// CFC twin of T_SafeTwoHand_Tests: the same tests drawn as CFC diagrams, the way a TwinSAFE project is authored.
    FUNCTION_BLOCK T_SafeTwoHand_Tests_CFC EXTENDS T_SafeCfcTestSuite
    VAR
    // Test_BothHandsGiveOutputAndReleaseNeedsBothOff
    group_1 : T_SafeGroup;
    fb_1 : T_SafeTwoHand(group := group_1);
    // Test_SecondHandWithoutFirstGivesTwoHandError
    group_2 : T_SafeGroup;
    fb_2 : T_SafeTwoHand(group := group_2);
    // Test_HandDiscrepancyTimeout
    group_3 : T_SafeGroup;
    // SafeInputsAfterDiscError TRUE (not the default) so the error waits for both hands released (diag bit 10)
    fb_3 : T_SafeTwoHand(group := group_3) := (Parameters := (HandDiscrepancyTime := T#100MS, SafeInputsAfterDiscError := TRUE));
    t0_3 : TON;
    t1_3 : TON;
    trig1_3 : R_TRIG;
END_VAR

Test_BothHandsGiveOutputAndReleaseNeedsBothOff();
Test_SecondHandWithoutFirstGivesTwoHandError();
Test_HandDiscrepancyTimeout();

METHOD PRIVATE Test_BothHandsGiveOutputAndReleaseNeedsBothOff
// note: this text did not pass the execution check against the stored diagram
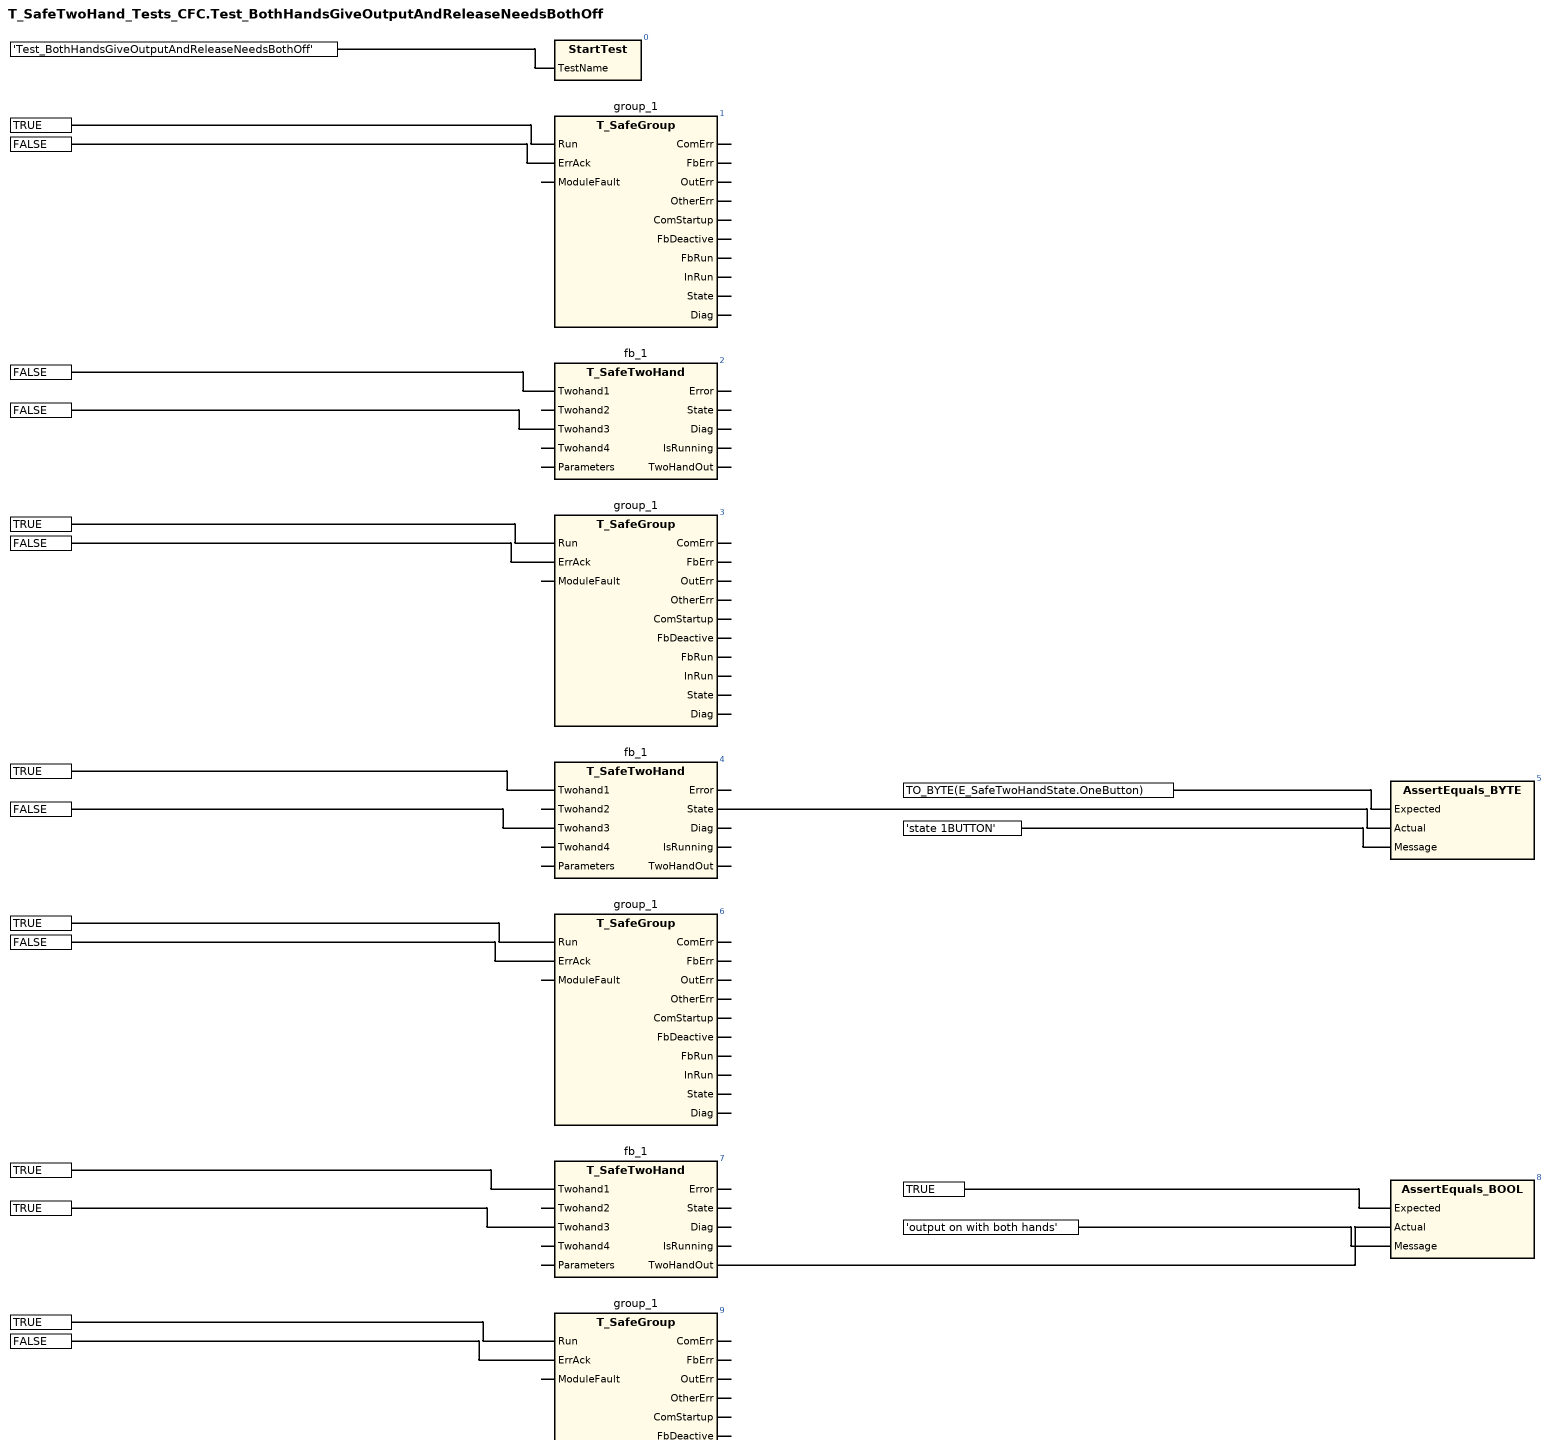
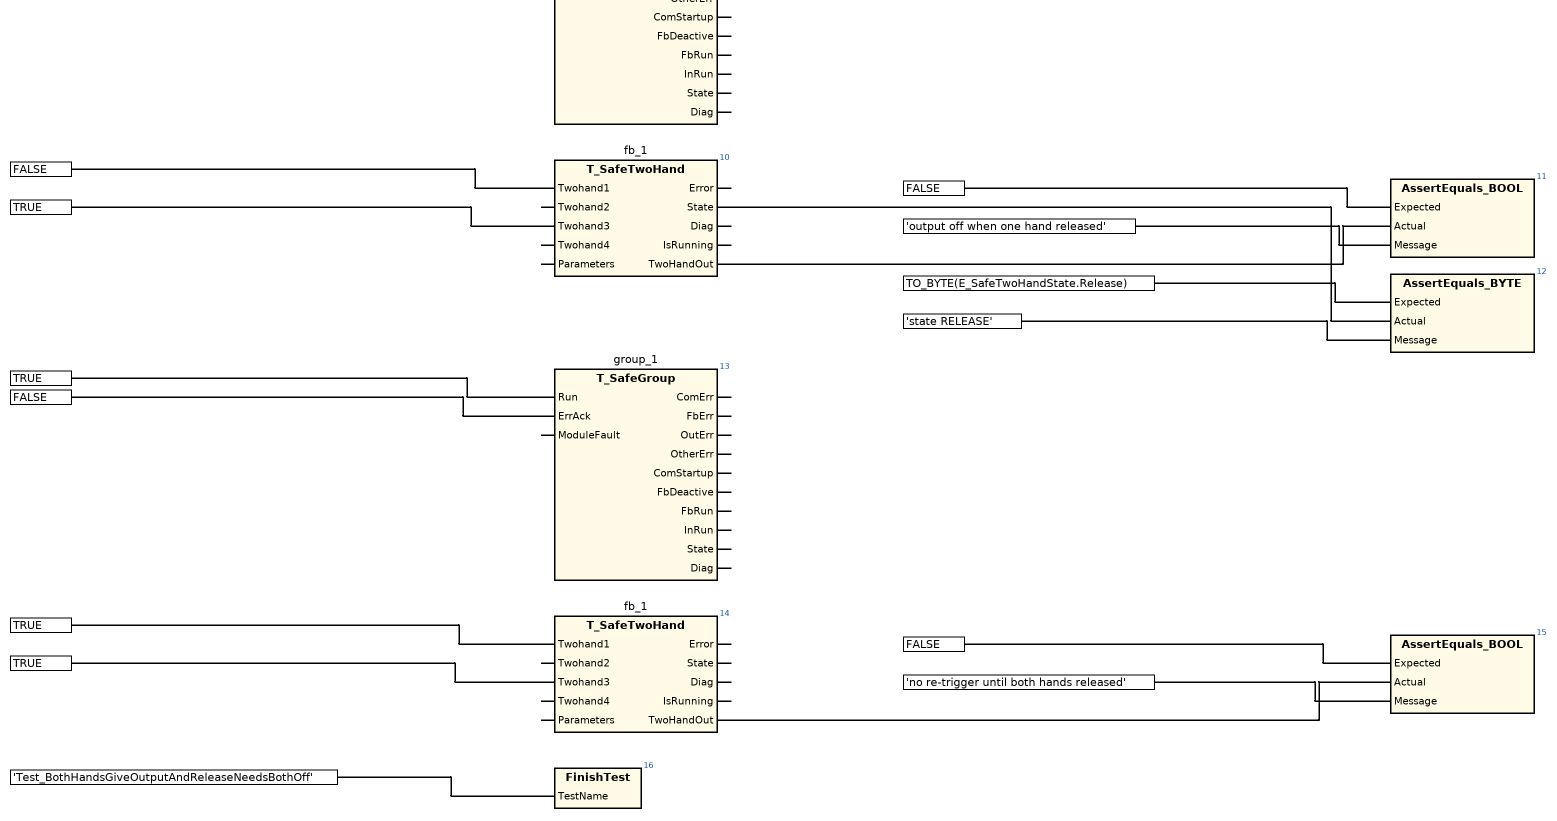
StartTest(TestName := 'Test_BothHandsGiveOutputAndReleaseNeedsBothOff');
group_1(Run := TRUE, ErrAck := FALSE); // T_SafeGroup
fb_1(Twohand1 := FALSE, Twohand3 := FALSE); // T_SafeTwoHand
group_1(Run := TRUE, ErrAck := FALSE); // T_SafeGroup
fb_1(Twohand1 := TRUE, Twohand3 := FALSE); // T_SafeTwoHand
AssertEquals_BYTE(Expected := TO_BYTE(E_SafeTwoHandState.OneButton), Actual := fb_1.State, Message := 'state 1BUTTON');
group_1(Run := TRUE, ErrAck := FALSE); // T_SafeGroup
fb_1(Twohand1 := TRUE, Twohand3 := TRUE); // T_SafeTwoHand
AssertEquals_BOOL(Expected := TRUE, Actual := fb_1.TwoHandOut, Message := 'output on with both hands');
group_1(Run := TRUE, ErrAck := FALSE); // T_SafeGroup
fb_1(Twohand1 := FALSE, Twohand3 := TRUE); // T_SafeTwoHand
AssertEquals_BOOL(Expected := FALSE, Actual := fb_1.TwoHandOut, Message := 'output off when one hand released');
AssertEquals_BYTE(Expected := TO_BYTE(E_SafeTwoHandState.Release), Actual := fb_1.State, Message := 'state RELEASE');
group_1(Run := TRUE, ErrAck := FALSE); // T_SafeGroup
fb_1(Twohand1 := TRUE, Twohand3 := TRUE); // T_SafeTwoHand
AssertEquals_BOOL(Expected := FALSE, Actual := fb_1.TwoHandOut, Message := 'no re-trigger until both hands released');
FinishTest(TestName := 'Test_BothHandsGiveOutputAndReleaseNeedsBothOff');
END_METHOD

METHOD PRIVATE Test_SecondHandWithoutFirstGivesTwoHandError
// note: this text did not pass the execution check against the stored diagram
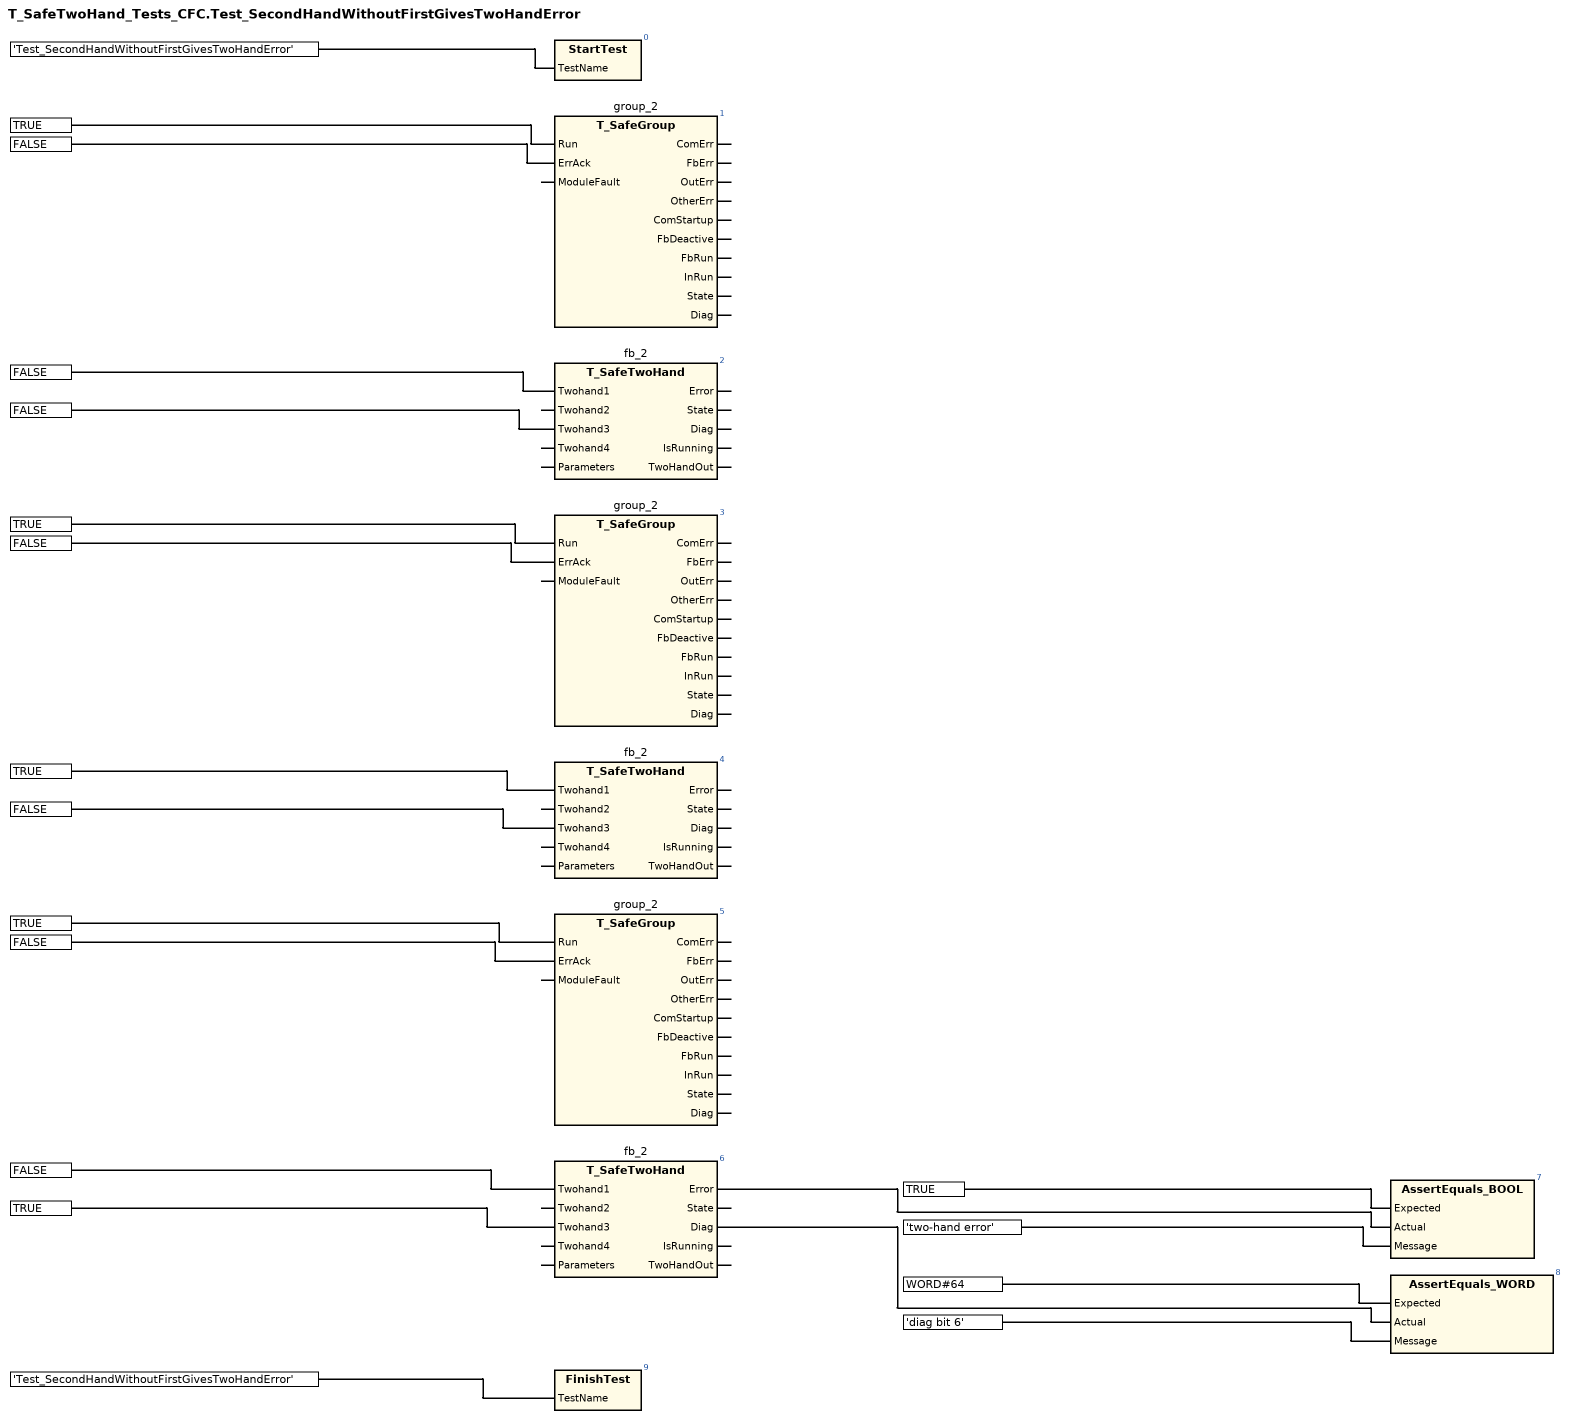
StartTest(TestName := 'Test_SecondHandWithoutFirstGivesTwoHandError');
group_2(Run := TRUE, ErrAck := FALSE); // T_SafeGroup
fb_2(Twohand1 := FALSE, Twohand3 := FALSE); // T_SafeTwoHand
group_2(Run := TRUE, ErrAck := FALSE); // T_SafeGroup
fb_2(Twohand1 := TRUE, Twohand3 := FALSE); // T_SafeTwoHand
group_2(Run := TRUE, ErrAck := FALSE); // T_SafeGroup
fb_2(Twohand1 := FALSE, Twohand3 := TRUE); // T_SafeTwoHand
AssertEquals_BOOL(Expected := TRUE, Actual := fb_2.Error, Message := 'two-hand error');
AssertEquals_WORD(Expected := WORD#64, Actual := fb_2.Diag, Message := 'diag bit 6');
FinishTest(TestName := 'Test_SecondHandWithoutFirstGivesTwoHandError');
END_METHOD

METHOD PRIVATE Test_HandDiscrepancyTimeout
// note: this text did not pass the execution check against the stored diagram
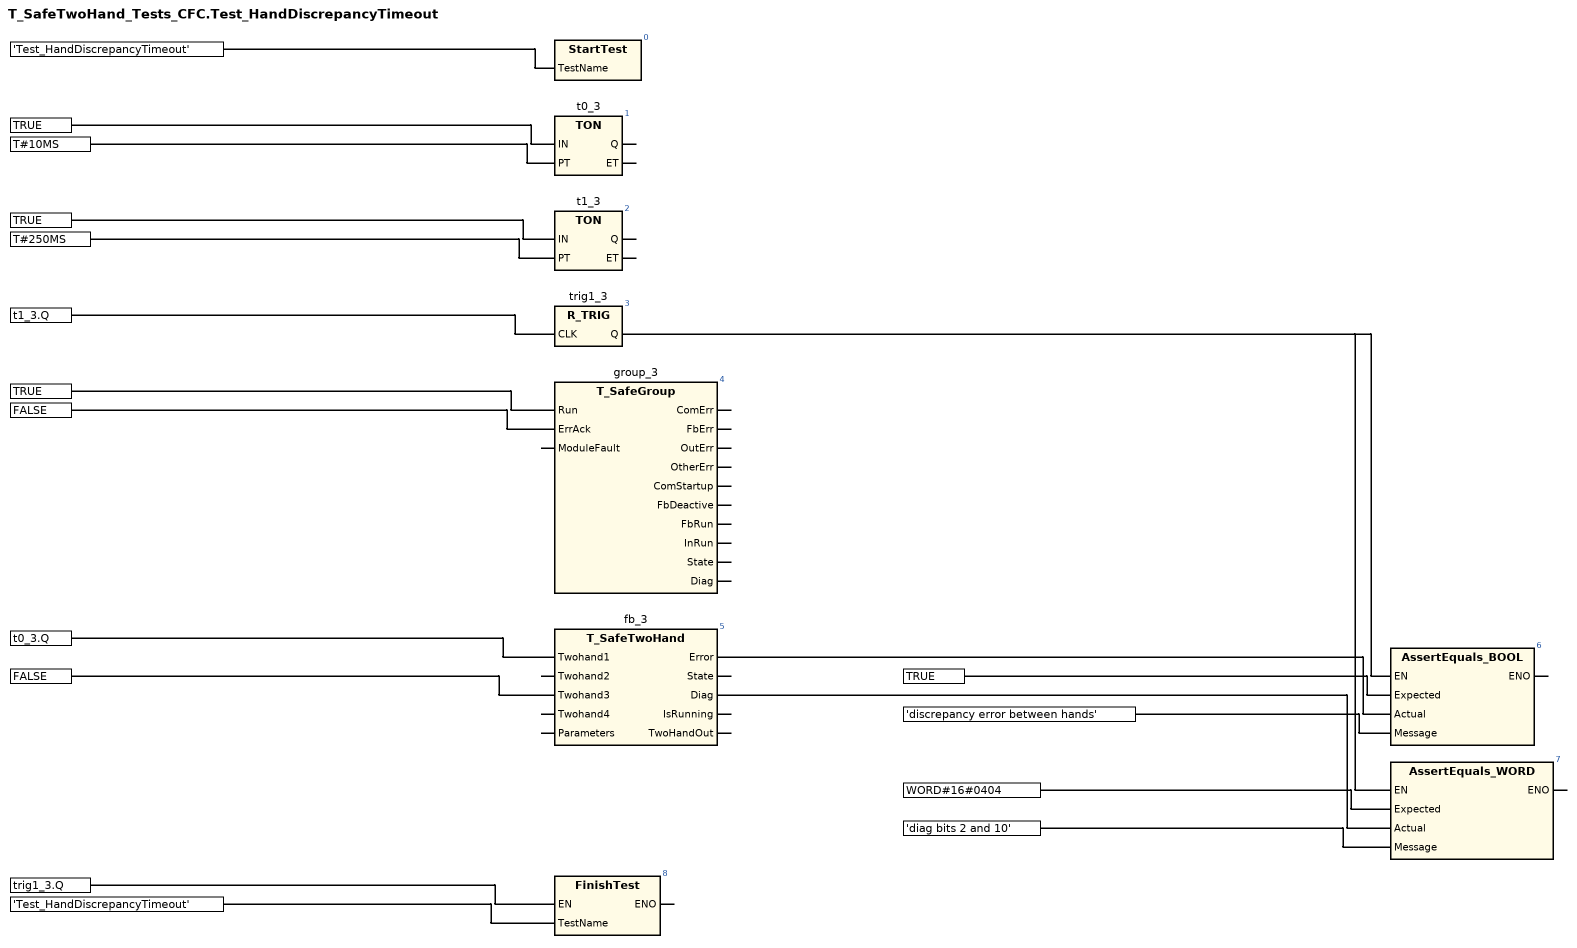
StartTest(TestName := 'Test_HandDiscrepancyTimeout');
t0_3(IN := TRUE, PT := T#10MS); // TON
t1_3(IN := TRUE, PT := T#250MS); // TON
trig1_3(CLK := t1_3.Q); // R_TRIG
group_3(Run := TRUE, ErrAck := FALSE); // T_SafeGroup
fb_3(Twohand1 := t0_3.Q, Twohand3 := FALSE); // T_SafeTwoHand
IF trig1_3.Q THEN AssertEquals_BOOL(Expected := TRUE, Actual := fb_3.Error, Message := 'discrepancy error between hands'); END_IF
IF trig1_3.Q THEN AssertEquals_WORD(Expected := WORD#16#0404, Actual := fb_3.Diag, Message := 'diag bits 2 and 10'); END_IF
IF trig1_3.Q THEN FinishTest(TestName := 'Test_HandDiscrepancyTimeout'); END_IF
END_METHOD

END_FUNCTION_BLOCK

(* stored: Version 1.1.0.1, ProductVersion 3.1.4026.22
   POU T_SafeTwoHand_Tests_CFC: Id {f7af8590-745c-5128-98b7-0cb820aa0a95}, SpecialFunc None
   Method Test_BothHandsGiveOutputAndReleaseNeedsBothOff: Id {58fb6d64-c76c-5eeb-80af-969a32e6bf17}
   Method Test_SecondHandWithoutFirstGivesTwoHandError: Id {85700aaf-46c4-58dc-b80a-494cba27532f}
   Method Test_HandDiscrepancyTimeout: Id {93ba127a-e4db-553e-be62-958c5a47c2b0} *)
